PROGRAM MAIN
VAR
	fbT1 : FB_IO_Test;
END_VAR

Tc3_PlcTestFramework.F_CallTestController();

END_PROGRAM

(* stored: Version 1.1.0.1
   POU MAIN: Id {adcb8fba-986a-4ac3-b18f-4d3d4a72882f}, SpecialFunc None *)
